(* IEC 61131-3 sources: repolevel_ST_code_completion/output/0121完整版本/repoeval_Proxy_Application/readful_result_before_fix, 2 files *)

(* ---- Proxy.st ---- *)
{attribute 'enable_dynamic_creation'}
FUNCTION_BLOCK Proxy IMPLEMENTS  Subject_Interface
VAR_INPUT
END_VAR
VAR_OUTPUT
END_VAR
VAR
	refToRealSubject : POINTER TO Realsubject;
	iTempPassword : INT;
END_VAR
VAR_STAT
	iRealPassword : INT := 1234;
END_VAR

METHOD fb_init
VAR_INPUT
	bInitRetains : BOOL;
	bInCopyCode : BOOL;
	ptrToRealSubject : POINTER TO Realsubject;
	iTempPassword : INT;
	iSetValue : INT;
	bReadWrite : BOOL;
END_VAR
VAR_OUTPUT
END_VAR
VAR
	refToRealSubject : POINTER TO Realsubject;
	iTempPassword : INT;
END_VAR

IF ptrToRealSubject <> 0 THEN
	refToRealSubject := ptrToRealSubject;
END_IF;

IF iTempPassword = iRealPassword THEN
	IF bReadWrite THEN
		refToRealSubject^.iProp := iSetValue;
	ELSE
		iSetValue := refToRealSubject^.iProp;
	END_IF;
END_IF;
END_FUNCTION_BLOCK

(* ---- Realsubject.st ---- *)
{attribute 'enable_dynamic_creation'}
FUNCTION_BLOCK Realsubject IMPLEMENTS  Subject_Interface
VAR_INPUT
END_VAR
VAR_OUTPUT
END_VAR
VAR
    // Variable to get and set values
    iProp: INT;
END_VAR

VAR_STAT
    // No static variables required for this implementation
END_VAR

METHOD PUBLIC Get_Method : INT
VAR
END_VAR
Get_Method := THIS^.iProp;

METHOD PUBLIC Set_Method
VAR_INPUT
    num : INT; // Value to be set on the iProp variable
END_VAR
THIS^.iProp := num;
END_FUNCTION_BLOCK
